TYPE "DT_REFERENCE_ALL"
VERSION : 0.1
   STRUCT
      WATER_LEVEL : "DT_REFERENCE_SOLO";
      WATER_PRESSURE : "DT_REFERENCE_SOLO";
      ACTIVE_POWER : "DT_REFERENCE_SOLO";
      OPENNESS : "DT_REFERENCE_SOLO";
      SPEED : "DT_REFERENCE_SOLO";
      KAPLAN_DISTRIBUTOR : "DT_REFERENCE_SOLO";
      KAPLAN_RUNNER : "DT_REFERENCE_SOLO";
      FRANCIS_DISTRIBUTOR : "DT_REFERENCE_SOLO";
      CROSS_FLOW_VALVE_1 : "DT_REFERENCE_SOLO";
      CROSS_FLOW_VALVE_2 : "DT_REFERENCE_SOLO";
      PELTON_DEFLECTOR : Array[1..6] of "DT_REFERENCE_SOLO";
      PELTON_NOZZLE : Array[1..6] of "DT_REFERENCE_SOLO";
      EXC_VOLTAGE : "DT_REFERENCE_SOLO";
      EXC_REACTIVE_POWER : "DT_REFERENCE_SOLO";
      EXC_POWER_FACTOR : "DT_REFERENCE_SOLO";
      Element_25 : "DT_REFERENCE_SOLO";
      Element_26 : "DT_REFERENCE_SOLO";
      Element_27 : "DT_REFERENCE_SOLO";
      Element_28 : "DT_REFERENCE_SOLO";
      Element_29 : "DT_REFERENCE_SOLO";
      Element_30 : "DT_REFERENCE_SOLO";
      Element_31 : "DT_REFERENCE_SOLO";
   END_STRUCT;

END_TYPE

